PROGRAM Main
  VAR
    b01_start : BOOL;
    b01_motor : BOOL;
    b01_permit : BOOL;
    b01_guard : BOOL;
    b02_a : BOOL;
    b02_out : BOOL;
    b02_b : BOOL;
    b02_c : BOOL;
    b02_e : BOOL;
    b06_run : BOOL;
    b06_lamp1 : BOOL;
    b06_lamp2 : BOOL;
    b06_lamp3 : BOOL;
    b07_cmd : BOOL;
    b07_latch : BOOL;
    b07_unlatch : BOOL;
    b07_rise : BOOL;
    b07_fall : BOOL;
    b11_conveyor_section_one_upstream_permissive_signal : BOOL;
    TON0 : TON;
    b11_conveyor_section_one_downstream_motor_run_command : BOOL;
    b11_conveyor_section_one_start_delay_preset_time_value : TIME;
    b11_conveyor_section_one_start_delay_elapsed_time_value : TIME;
  END_VAR
  VAR  (* added by the conversion: wires and edge detectors of the diagram *)
    R_TRIG1 : R_TRIG;
    F_TRIG2 : F_TRIG;
  END_VAR

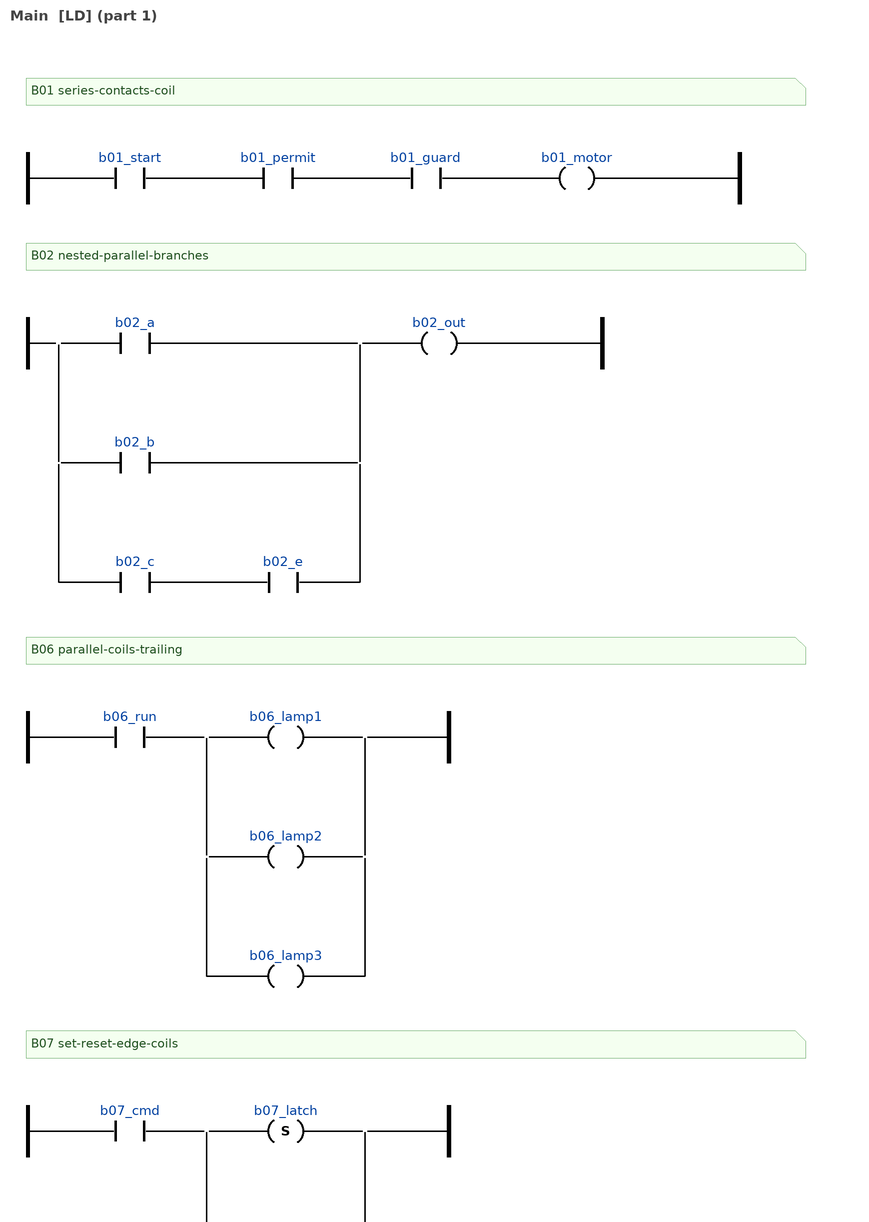
(* LD diagram, written out as Structured Text *)
(* B01 series-contacts-coil *)
b01_motor := b01_start AND b01_permit AND b01_guard;
(* B02 nested-parallel-branches *)
b02_out := b02_a OR b02_b OR b02_c AND b02_e;
(* B06 parallel-coils-trailing *)
b06_lamp1 := b06_run;
b06_lamp2 := b06_run;
b06_lamp3 := b06_run;
(* B07 set-reset-edge-coils *)
IF b07_cmd THEN b07_latch := TRUE; END_IF;
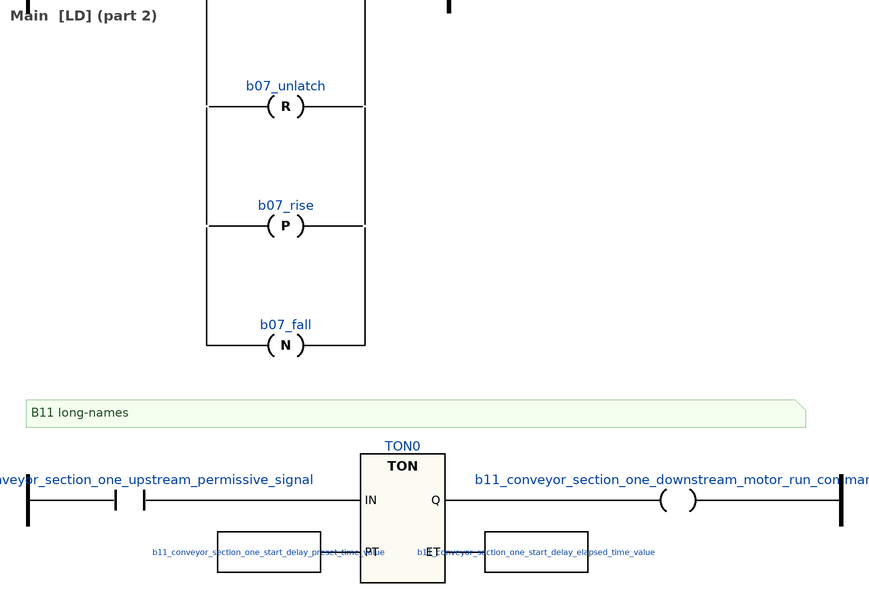
IF b07_cmd THEN b07_unlatch := FALSE; END_IF;
R_TRIG1(CLK := b07_cmd);
b07_rise := R_TRIG1.Q;
F_TRIG2(CLK := b07_cmd);
b07_fall := F_TRIG2.Q;
(* B11 long-names *)
TON0(IN := b11_conveyor_section_one_upstream_permissive_signal, PT := b11_conveyor_section_one_start_delay_preset_time_value);
b11_conveyor_section_one_downstream_motor_run_command := TON0.Q;
b11_conveyor_section_one_start_delay_elapsed_time_value := TON0.ET;
END_PROGRAM
